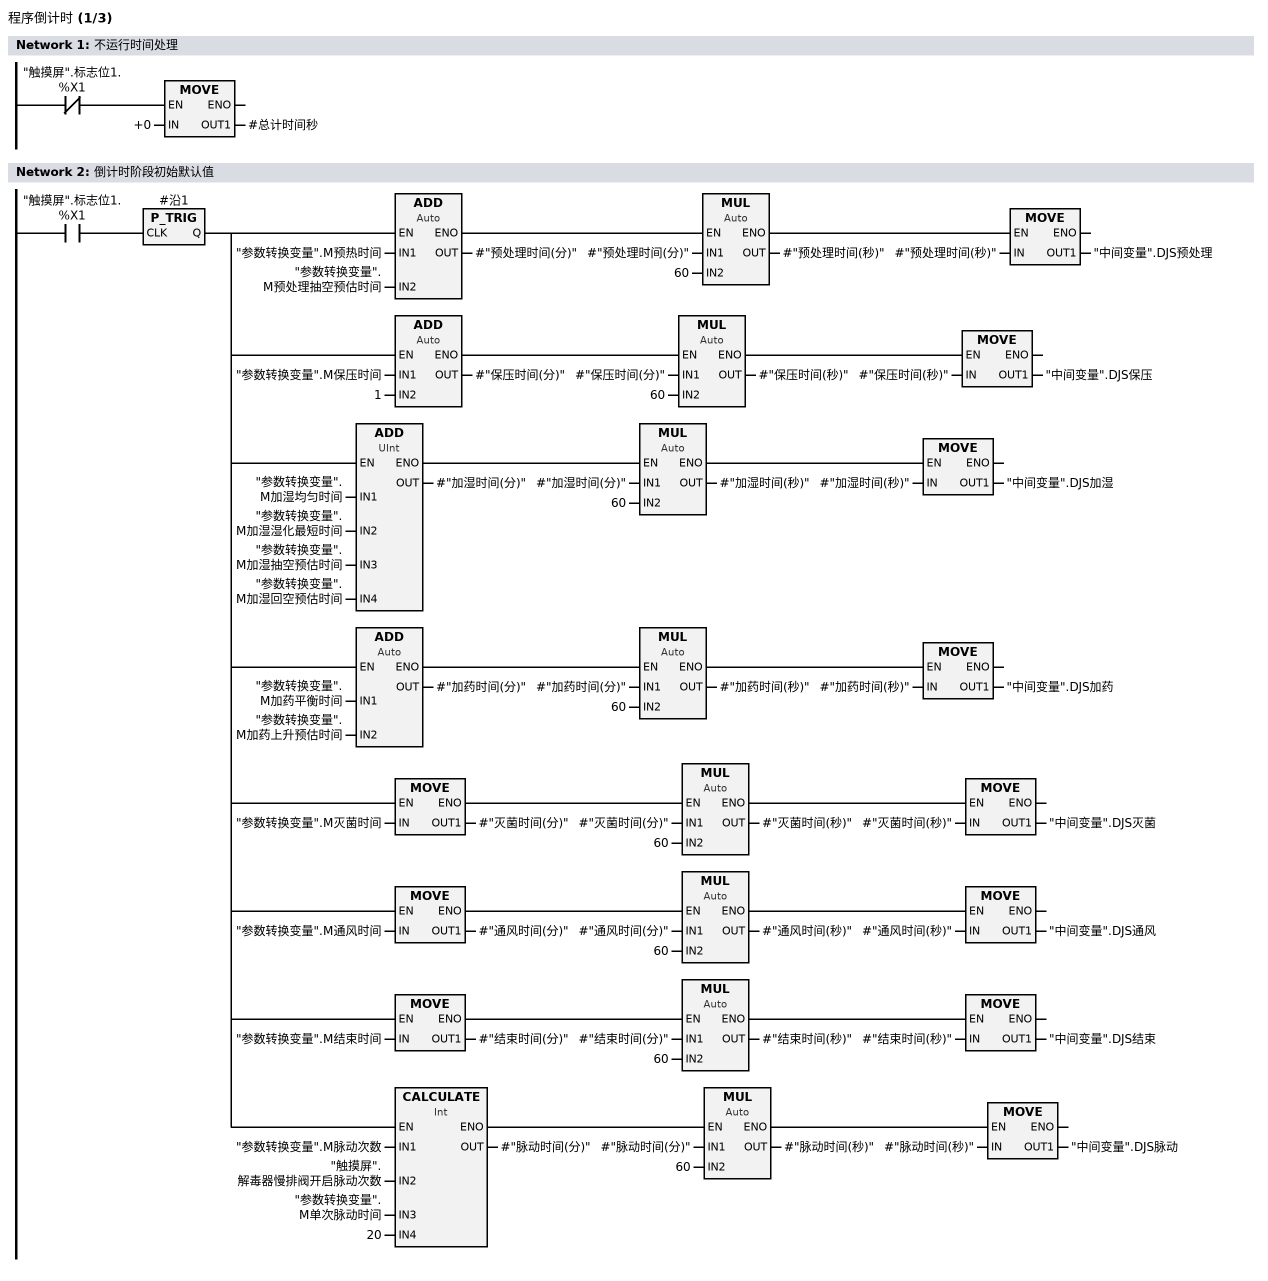
   RUNG wire#powerrail
      I_Contact( "触摸屏".标志位1.%X1 )
      Move(in := +0, out1 => #总计时间秒)
   END_RUNG
   // the same network as SCL:
   IF NOT "触摸屏".标志位1.%X1 THEN #总计时间秒 := +0; END_IF;
END_REGION

REGION Network 2: 倒计时阶段初始默认值
   RUNG wire#powerrail
      Contact( "触摸屏".标志位1.%X1 )
      P_Trig( #沿1 )
      wire#w1
      Add(in1 := "参数转换变量".M预热时间, in2 := "参数转换变量".M预处理抽空预估时间, out => #"预处理时间(分)")
      Mul(in1 := #"预处理时间(分)", in2 := 60, out => #"预处理时间(秒)")
      Move(in := #"预处理时间(秒)", out1 => "中间变量".DJS预处理)
   END_RUNG
   RUNG wire#w1
      Add(in1 := "参数转换变量".M保压时间, in2 := 1, out => #"保压时间(分)")
      Mul(in1 := #"保压时间(分)", in2 := 60, out => #"保压时间(秒)")
      Move(in := #"保压时间(秒)", out1 => "中间变量".DJS保压)
   END_RUNG
   RUNG wire#w1
      { S7_Templates := "SrcType := UInt" } Add(in1 := "参数转换变量".M加湿均匀时间, in2 := "参数转换变量".M加湿湿化最短时间, in3 := "参数转换变量".M加湿抽空预估时间, in4 := "参数转换变量".M加湿回空预估时间, out => #"加湿时间(分)")
      Mul(in1 := #"加湿时间(分)", in2 := 60, out => #"加湿时间(秒)")
      Move(in := #"加湿时间(秒)", out1 => "中间变量".DJS加湿)
   END_RUNG
   RUNG wire#w1
      Add(in1 := "参数转换变量".M加药平衡时间, in2 := "参数转换变量".M加药上升预估时间, out => #"加药时间(分)")
      Mul(in1 := #"加药时间(分)", in2 := 60, out => #"加药时间(秒)")
      Move(in := #"加药时间(秒)", out1 => "中间变量".DJS加药)
   END_RUNG
   RUNG wire#w1
      Move(in := "参数转换变量".M灭菌时间, out1 => #"灭菌时间(分)")
      Mul(in1 := #"灭菌时间(分)", in2 := 60, out => #"灭菌时间(秒)")
      Move(in := #"灭菌时间(秒)", out1 => "中间变量".DJS灭菌)
   END_RUNG
   RUNG wire#w1
      Move(in := "参数转换变量".M通风时间, out1 => #"通风时间(分)")
      Mul(in1 := #"通风时间(分)", in2 := 60, out => #"通风时间(秒)")
      Move(in := #"通风时间(秒)", out1 => "中间变量".DJS通风)
   END_RUNG
   RUNG wire#w1
      Move(in := "参数转换变量".M结束时间, out1 => #"结束时间(分)")
      Mul(in1 := #"结束时间(分)", in2 := 60, out => #"结束时间(秒)")
      Move(in := #"结束时间(秒)", out1 => "中间变量".DJS结束)
   END_RUNG
   RUNG wire#w1
      { S7_Templates := "SrcType := Int"; S7_Expression := "(IN1-IN2)*IN3+IN2*IN4" } Calculate(in1 := "参数转换变量".M脉动次数, in2 := "触摸屏".解毒器慢排阀开启脉动次数, in3 := "参数转换变量".M单次脉动时间, in4 := 20, out => #"脉动时间(分)")
      Mul(in1 := #"脉动时间(分)", in2 := 60, out => #"脉动时间(秒)")
      Move(in := #"脉动时间(秒)", out1 => "中间变量".DJS脉动)
   END_RUNG
   // the same network as SCL:
   #_w1 := "触摸屏".标志位1.%X1 AND NOT #沿1;   // rising edge
   #沿1 := "触摸屏".标志位1.%X1;
   IF #_w1 THEN
       #"预处理时间(分)" := "参数转换变量".M预热时间 + "参数转换变量".M预处理抽空预估时间;
       #"预处理时间(秒)" := #"预处理时间(分)" * 60;
       "中间变量".DJS预处理 := #"预处理时间(秒)";
       #"保压时间(分)" := "参数转换变量".M保压时间 + 1;
       #"保压时间(秒)" := #"保压时间(分)" * 60;
       "中间变量".DJS保压 := #"保压时间(秒)";
       #"加湿时间(分)" := "参数转换变量".M加湿均匀时间 + "参数转换变量".M加湿湿化最短时间 + "参数转换变量".M加湿抽空预估时间 + "参数转换变量".M加湿回空预估时间;
       #"加湿时间(秒)" := #"加湿时间(分)" * 60;
       "中间变量".DJS加湿 := #"加湿时间(秒)";
       #"加药时间(分)" := "参数转换变量".M加药平衡时间 + "参数转换变量".M加药上升预估时间;
       #"加药时间(秒)" := #"加药时间(分)" * 60;
       "中间变量".DJS加药 := #"加药时间(秒)";
       #"灭菌时间(分)" := "参数转换变量".M灭菌时间;
       #"灭菌时间(秒)" := #"灭菌时间(分)" * 60;
       "中间变量".DJS灭菌 := #"灭菌时间(秒)";
       #"通风时间(分)" := "参数转换变量".M通风时间;
       #"通风时间(秒)" := #"通风时间(分)" * 60;
       "中间变量".DJS通风 := #"通风时间(秒)";
       #"结束时间(分)" := "参数转换变量".M结束时间;
       #"结束时间(秒)" := #"结束时间(分)" * 60;
       "中间变量".DJS结束 := #"结束时间(秒)";
       #"脉动时间(分)" := ("参数转换变量".M脉动次数-"触摸屏".解毒器慢排阀开启脉动次数)*"参数转换变量".M单次脉动时间+"触摸屏".解毒器慢排阀开启脉动次数*20;
       #"脉动时间(秒)" := #"脉动时间(分)" * 60;
       "中间变量".DJS脉动 := #"脉动时间(秒)";
   END_IF;
END_REGION

REGION Network 3: 倒计时
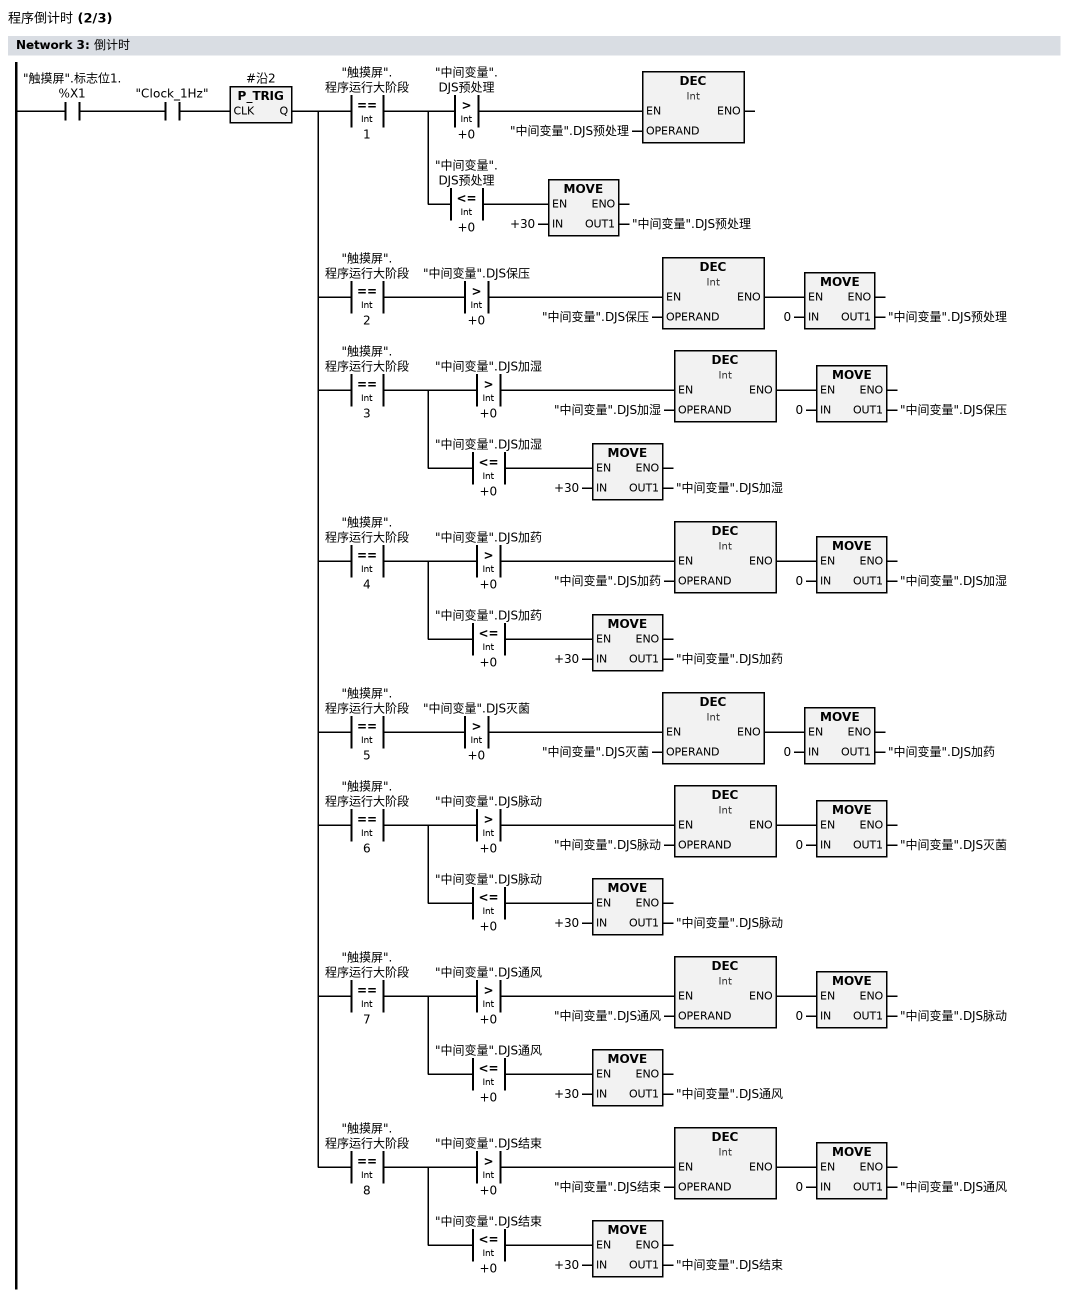
   RUNG wire#powerrail
      Contact( "触摸屏".标志位1.%X1 )
      Contact( "Clock_1Hz" )
      P_Trig( #沿2 )
      wire#w1
      { S7_Templates := "SrcType := Int" } EQ_Contact(in1 := "触摸屏".程序运行大阶段, in2 := 1)
      wire#w2
      { S7_Templates := "SrcType := Int" } GT_Contact(in1 := "中间变量".DJS预处理, in2 := +0)
      { S7_Templates := "DestType := Int" } Dec( "中间变量".DJS预处理 )
   END_RUNG
   RUNG wire#w2
      { S7_Templates := "SrcType := Int" } LE_Contact(in1 := "中间变量".DJS预处理, in2 := +0)
      Move(in := +30, out1 => "中间变量".DJS预处理)
   END_RUNG
   RUNG wire#w1
      { S7_Templates := "SrcType := Int" } EQ_Contact(in1 := "触摸屏".程序运行大阶段, in2 := 2)
      { S7_Templates := "SrcType := Int" } GT_Contact(in1 := "中间变量".DJS保压, in2 := +0)
      { S7_Templates := "DestType := Int" } Dec( "中间变量".DJS保压 )
      Move(in := 0, out1 => "中间变量".DJS预处理)
   END_RUNG
   RUNG wire#w1
      { S7_Templates := "SrcType := Int" } EQ_Contact(in1 := "触摸屏".程序运行大阶段, in2 := 3)
      wire#w3
      { S7_Templates := "SrcType := Int" } GT_Contact(in1 := "中间变量".DJS加湿, in2 := +0)
      { S7_Templates := "DestType := Int" } Dec( "中间变量".DJS加湿 )
      Move(in := 0, out1 => "中间变量".DJS保压)
   END_RUNG
   RUNG wire#w3
      { S7_Templates := "SrcType := Int" } LE_Contact(in1 := "中间变量".DJS加湿, in2 := +0)
      Move(in := +30, out1 => "中间变量".DJS加湿)
   END_RUNG
   RUNG wire#w1
      { S7_Templates := "SrcType := Int" } EQ_Contact(in1 := "触摸屏".程序运行大阶段, in2 := 4)
      wire#w4
      { S7_Templates := "SrcType := Int" } GT_Contact(in1 := "中间变量".DJS加药, in2 := +0)
      { S7_Templates := "DestType := Int" } Dec( "中间变量".DJS加药 )
      Move(in := 0, out1 => "中间变量".DJS加湿)
   END_RUNG
   RUNG wire#w4
      { S7_Templates := "SrcType := Int" } LE_Contact(in1 := "中间变量".DJS加药, in2 := +0)
      Move(in := +30, out1 => "中间变量".DJS加药)
   END_RUNG
   RUNG wire#w1
      { S7_Templates := "SrcType := Int" } EQ_Contact(in1 := "触摸屏".程序运行大阶段, in2 := 5)
      { S7_Templates := "SrcType := Int" } GT_Contact(in1 := "中间变量".DJS灭菌, in2 := +0)
      { S7_Templates := "DestType := Int" } Dec( "中间变量".DJS灭菌 )
      Move(in := 0, out1 => "中间变量".DJS加药)
   END_RUNG
   RUNG wire#w1
      { S7_Templates := "SrcType := Int" } EQ_Contact(in1 := "触摸屏".程序运行大阶段, in2 := 6)
      wire#w5
      { S7_Templates := "SrcType := Int" } GT_Contact(in1 := "中间变量".DJS脉动, in2 := +0)
      { S7_Templates := "DestType := Int" } Dec( "中间变量".DJS脉动 )
      Move(in := 0, out1 => "中间变量".DJS灭菌)
   END_RUNG
   RUNG wire#w5
      { S7_Templates := "SrcType := Int" } LE_Contact(in1 := "中间变量".DJS脉动, in2 := +0)
      Move(in := +30, out1 => "中间变量".DJS脉动)
   END_RUNG
   RUNG wire#w1
      { S7_Templates := "SrcType := Int" } EQ_Contact(in1 := "触摸屏".程序运行大阶段, in2 := 7)
      wire#w6
      { S7_Templates := "SrcType := Int" } GT_Contact(in1 := "中间变量".DJS通风, in2 := +0)
      { S7_Templates := "DestType := Int" } Dec( "中间变量".DJS通风 )
      Move(in := 0, out1 => "中间变量".DJS脉动)
   END_RUNG
   RUNG wire#w6
      { S7_Templates := "SrcType := Int" } LE_Contact(in1 := "中间变量".DJS通风, in2 := +0)
      Move(in := +30, out1 => "中间变量".DJS通风)
   END_RUNG
   RUNG wire#w1
      { S7_Templates := "SrcType := Int" } EQ_Contact(in1 := "触摸屏".程序运行大阶段, in2 := 8)
      wire#w7
      { S7_Templates := "SrcType := Int" } GT_Contact(in1 := "中间变量".DJS结束, in2 := +0)
      { S7_Templates := "DestType := Int" } Dec( "中间变量".DJS结束 )
      Move(in := 0, out1 => "中间变量".DJS通风)
   END_RUNG
   RUNG wire#w7
      { S7_Templates := "SrcType := Int" } LE_Contact(in1 := "中间变量".DJS结束, in2 := +0)
      Move(in := +30, out1 => "中间变量".DJS结束)
   END_RUNG
   // the same network as SCL:
   #_w1 := "触摸屏".标志位1.%X1 AND "Clock_1Hz";
   #_w2 := #_w1 AND NOT #沿2;   // rising edge
   #沿2 := #_w1;
   #_w3 := #_w2 AND ("触摸屏".程序运行大阶段 = 1);
   IF #_w3 AND ("中间变量".DJS预处理 > +0) THEN "中间变量".DJS预处理 := "中间变量".DJS预处理 - 1; END_IF;
   IF #_w3 AND ("中间变量".DJS预处理 <= +0) THEN "中间变量".DJS预处理 := +30; END_IF;
   #_w4 := #_w2 AND ("触摸屏".程序运行大阶段 = 2) AND ("中间变量".DJS保压 > +0);
   IF #_w4 THEN
       "中间变量".DJS保压 := "中间变量".DJS保压 - 1;
       "中间变量".DJS预处理 := 0;
   END_IF;
   #_w5 := #_w2 AND ("触摸屏".程序运行大阶段 = 3);
   #_w6 := #_w5 AND ("中间变量".DJS加湿 > +0);
   IF #_w6 THEN
       "中间变量".DJS加湿 := "中间变量".DJS加湿 - 1;
       "中间变量".DJS保压 := 0;
   END_IF;
   IF #_w5 AND ("中间变量".DJS加湿 <= +0) THEN "中间变量".DJS加湿 := +30; END_IF;
   #_w7 := #_w2 AND ("触摸屏".程序运行大阶段 = 4);
   #_w8 := #_w7 AND ("中间变量".DJS加药 > +0);
   IF #_w8 THEN
       "中间变量".DJS加药 := "中间变量".DJS加药 - 1;
       "中间变量".DJS加湿 := 0;
   END_IF;
   IF #_w7 AND ("中间变量".DJS加药 <= +0) THEN "中间变量".DJS加药 := +30; END_IF;
   #_w9 := #_w2 AND ("触摸屏".程序运行大阶段 = 5) AND ("中间变量".DJS灭菌 > +0);
   IF #_w9 THEN
       "中间变量".DJS灭菌 := "中间变量".DJS灭菌 - 1;
       "中间变量".DJS加药 := 0;
   END_IF;
   #_w10 := #_w2 AND ("触摸屏".程序运行大阶段 = 6);
   #_w11 := #_w10 AND ("中间变量".DJS脉动 > +0);
   IF #_w11 THEN
       "中间变量".DJS脉动 := "中间变量".DJS脉动 - 1;
       "中间变量".DJS灭菌 := 0;
   END_IF;
   IF #_w10 AND ("中间变量".DJS脉动 <= +0) THEN "中间变量".DJS脉动 := +30; END_IF;
   #_w12 := #_w2 AND ("触摸屏".程序运行大阶段 = 7);
   #_w13 := #_w12 AND ("中间变量".DJS通风 > +0);
   IF #_w13 THEN
       "中间变量".DJS通风 := "中间变量".DJS通风 - 1;
       "中间变量".DJS脉动 := 0;
   END_IF;
   IF #_w12 AND ("中间变量".DJS通风 <= +0) THEN "中间变量".DJS通风 := +30; END_IF;
   #_w14 := #_w2 AND ("触摸屏".程序运行大阶段 = 8);
   #_w15 := #_w14 AND ("中间变量".DJS结束 > +0);
   IF #_w15 THEN
       "中间变量".DJS结束 := "中间变量".DJS结束 - 1;
       "中间变量".DJS通风 := 0;
   END_IF;
   IF #_w14 AND ("中间变量".DJS结束 <= +0) THEN "中间变量".DJS结束 := +30; END_IF;
END_REGION

REGION Network 4: 阶段时间累加
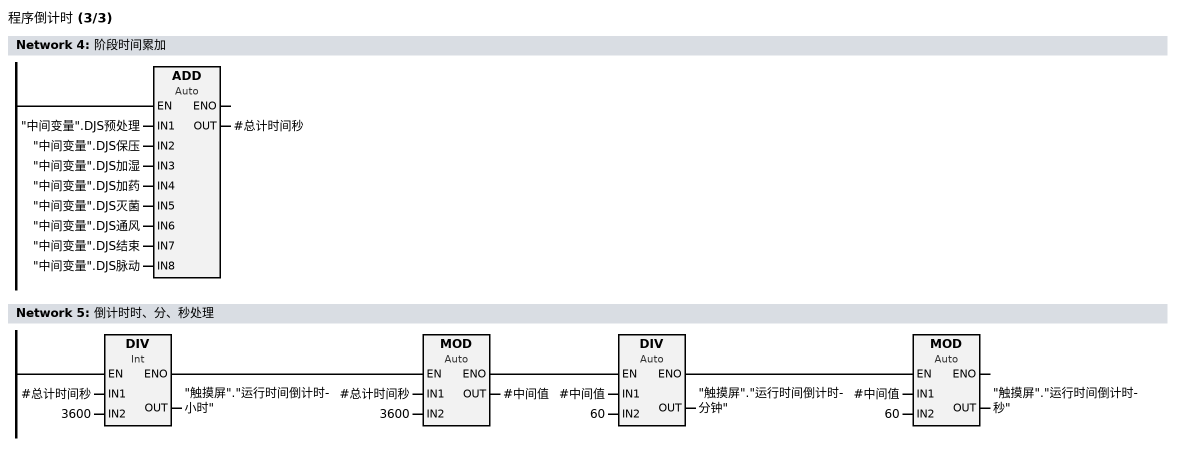
   RUNG wire#powerrail
      Add(in1 := "中间变量".DJS预处理, in2 := "中间变量".DJS保压, in3 := "中间变量".DJS加湿, in4 := "中间变量".DJS加药, in5 := "中间变量".DJS灭菌, in6 := "中间变量".DJS通风, in7 := "中间变量".DJS结束, in8 := "中间变量".DJS脉动, out => #总计时间秒)
   END_RUNG
   // the same network as SCL:
   #总计时间秒 := "中间变量".DJS预处理 + "中间变量".DJS保压 + "中间变量".DJS加湿 + "中间变量".DJS加药 + "中间变量".DJS灭菌 + "中间变量".DJS通风 + "中间变量".DJS结束 + "中间变量".DJS脉动;
END_REGION

REGION Network 5: 倒计时时、分、秒处理
   RUNG wire#powerrail
      { S7_Templates := "SrcType := Int" } Div(in1 := #总计时间秒, in2 := 3600, out => "触摸屏"."运行时间倒计时-小时")
      Mod(in1 := #总计时间秒, in2 := 3600, out => #中间值)
      Div(in1 := #中间值, in2 := 60, out => "触摸屏"."运行时间倒计时-分钟")
      Mod(in1 := #中间值, in2 := 60, out => "触摸屏"."运行时间倒计时-秒")
   END_RUNG
   // the same network as SCL:
   "触摸屏"."运行时间倒计时-小时" := #总计时间秒 / 3600;
   #中间值 := #总计时间秒 MOD 3600;
   "触摸屏"."运行时间倒计时-分钟" := #中间值 / 60;
   "触摸屏"."运行时间倒计时-秒" := #中间值 MOD 60;
END_REGION
END_FUNCTION_BLOCK

FUNCTION "计算倒计时" : Void   // FC6, LAD
{ S7_Optimized_Access := 'TRUE' }
VERSION : 0.1
   VAR_INPUT
      程序运行大阶段 : Int;
   END_VAR
   VAR_OUTPUT
      倒计时总秒数 : DInt;
      各阶段运行时间秒 : DInt;
      循环计数 : Int;
   END_VAR
   VAR_TEMP
      获取当前预制区阶段预估时间秒 : Int;
   END_VAR
BEGIN

REGION Network 1
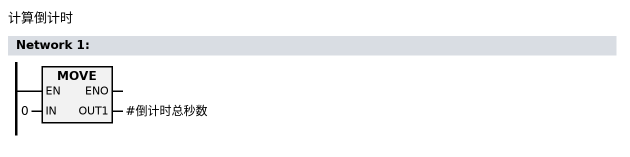
   RUNG wire#powerrail
      Move(in := 0, out1 => #倒计时总秒数)
   END_RUNG
   // the same network as SCL:
   #倒计时总秒数 := 0;
END_REGION

REGION Network 2 (SCL)
   IF #程序运行大阶段 >=0 AND #程序运行大阶段<=10  THEN
       FOR #循环计数 := #程序运行大阶段 TO 10 DO
           IF (#程序运行大阶段 < 8 OR #程序运行大阶段 > 9) THEN

               IF (#循环计数 <> 8 AND #循环计数 <> 9) THEN
                   "获取各阶段预估运行时间秒"(当前阶段名称 := #循环计数,
                                  当前阶段预估时间秒 => #各阶段运行时间秒);
               ELSE
                   #各阶段运行时间秒 := 0;

               END_IF;
           ELSE
               "获取各阶段预估运行时间秒"(当前阶段名称 := #循环计数,
                              当前阶段预估时间秒 => #各阶段运行时间秒);


           END_IF;
           #倒计时总秒数 := #倒计时总秒数 + #各阶段运行时间秒;


       END_FOR;

       END_IF;
END_REGION
END_FUNCTION

FUNCTION "获取各阶段预估运行时间秒" : Void   // FC18, LAD
{ S7_Optimized_Access := 'TRUE' }
VERSION : 0.1
   VAR_INPUT
      当前阶段名称 : Int;
   END_VAR
   VAR_OUTPUT
      当前阶段预估时间秒 : DInt;
   END_VAR
   VAR_TEMP
      沿1 : Bool;
      沿2 : Bool;
   END_VAR
   VAR_TEMP   // added for the SCL form of the ladder/FBD networks
      _w1 : Bool;
   END_VAR
BEGIN

REGION Network 1
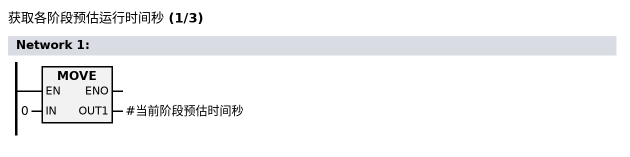
   RUNG wire#powerrail
      Move(in := 0, out1 => #当前阶段预估时间秒)
   END_RUNG
   // the same network as SCL:
   #当前阶段预估时间秒 := 0;
END_REGION

REGION Network 2: 倒计时阶段初始默认值
   // "触摸屏".程序类型.%X2:药罐处理、"触摸屏".程序类型.%X3:泄漏测试
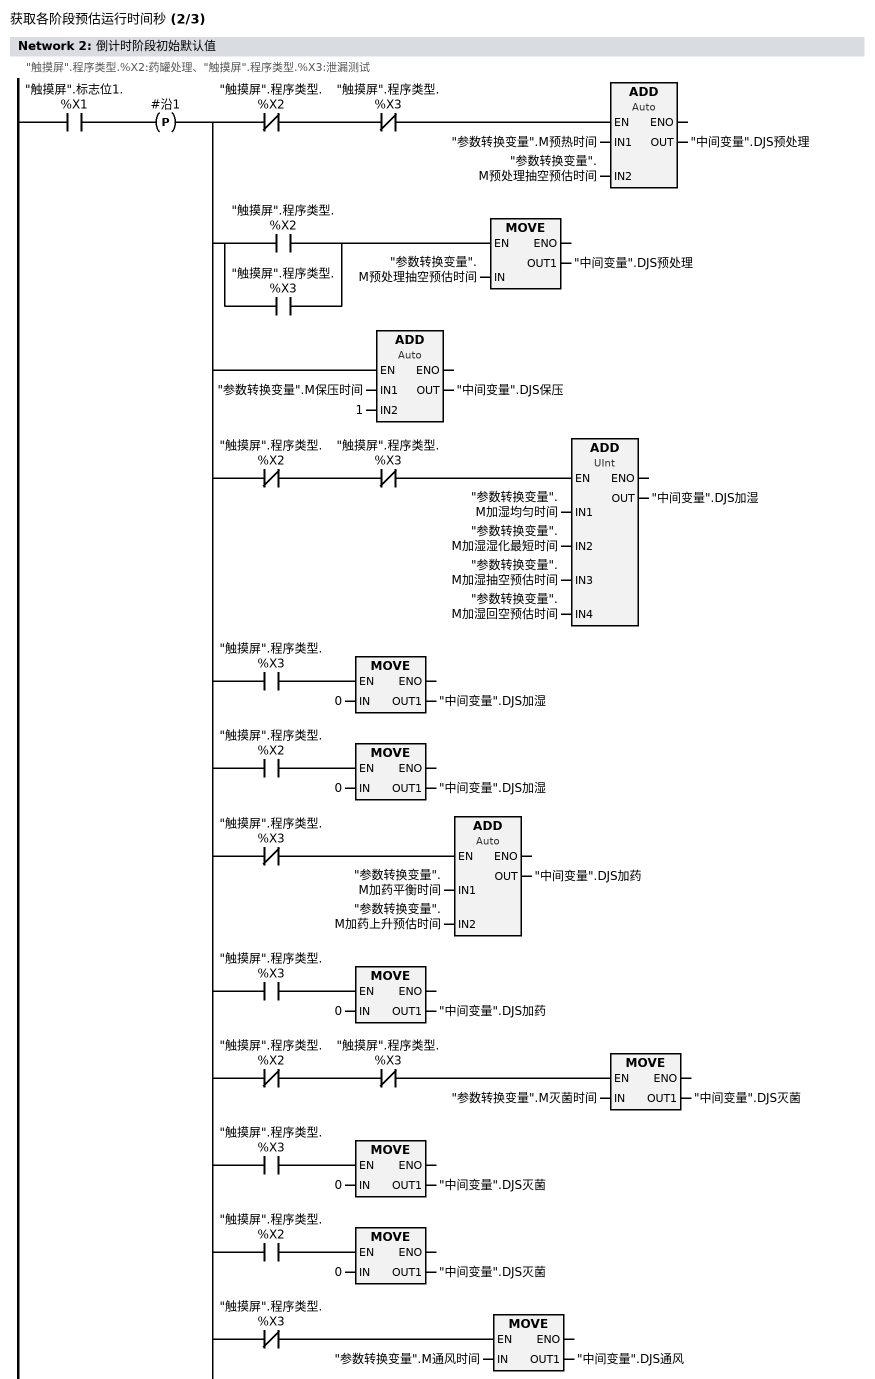
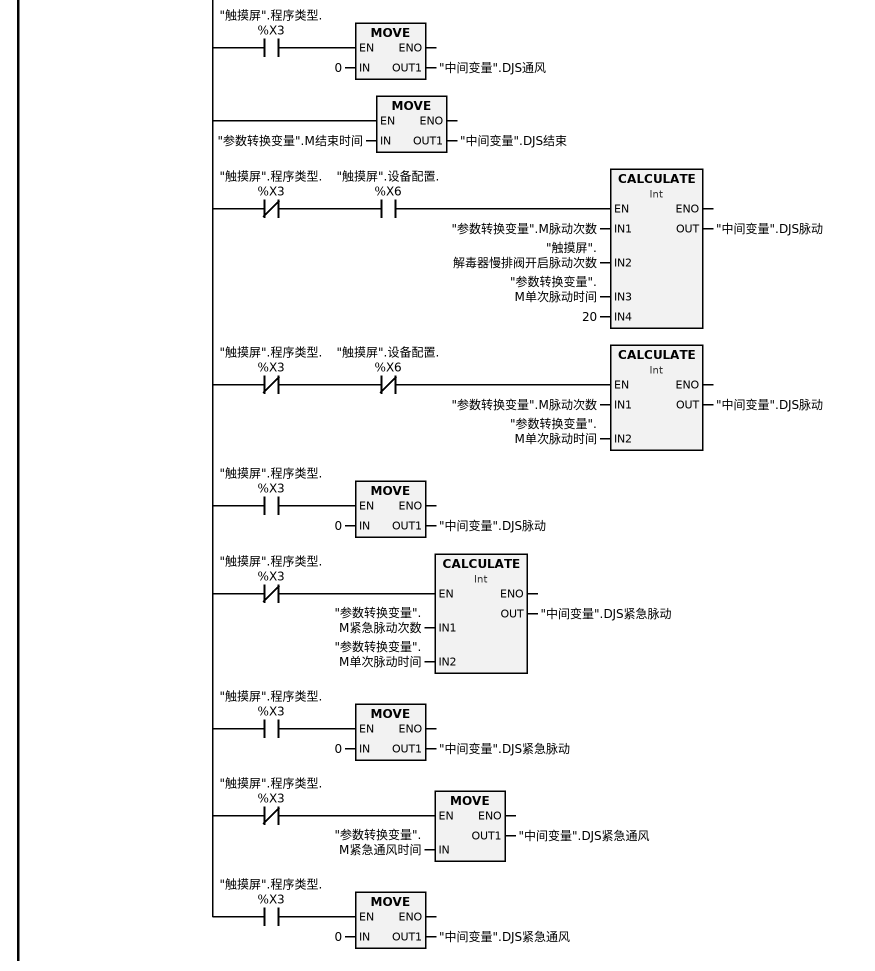
   RUNG wire#powerrail
      Contact( "触摸屏".标志位1.%X1 )
      P_Trig( #沿1 )
      wire#w1
      I_Contact( "触摸屏".程序类型.%X2 )
      I_Contact( "触摸屏".程序类型.%X3 )
      Add(in1 := "参数转换变量".M预热时间, in2 := "参数转换变量".M预处理抽空预估时间, out => "中间变量".DJS预处理)
   END_RUNG
   RUNG wire#w1
      Contact( "触摸屏".程序类型.%X2 )
      wire#w2
      Move(in := "参数转换变量".M预处理抽空预估时间, out1 => "中间变量".DJS预处理)
   END_RUNG
   RUNG wire#w1
      Contact( "触摸屏".程序类型.%X3 )
   END_RUNG wire#w2
   RUNG wire#w1
      Add(in1 := "参数转换变量".M保压时间, in2 := 1, out => "中间变量".DJS保压)
   END_RUNG
   RUNG wire#w1
      I_Contact( "触摸屏".程序类型.%X2 )
      I_Contact( "触摸屏".程序类型.%X3 )
      { S7_Templates := "SrcType := UInt" } Add(in1 := "参数转换变量".M加湿均匀时间, in2 := "参数转换变量".M加湿湿化最短时间, in3 := "参数转换变量".M加湿抽空预估时间, in4 := "参数转换变量".M加湿回空预估时间, out => "中间变量".DJS加湿)
   END_RUNG
   RUNG wire#w1
      Contact( "触摸屏".程序类型.%X3 )
      Move(in := 0, out1 => "中间变量".DJS加湿)
   END_RUNG
   RUNG wire#w1
      Contact( "触摸屏".程序类型.%X2 )
      Move(in := 0, out1 => "中间变量".DJS加湿)
   END_RUNG
   RUNG wire#w1
      I_Contact( "触摸屏".程序类型.%X3 )
      Add(in1 := "参数转换变量".M加药平衡时间, in2 := "参数转换变量".M加药上升预估时间, out => "中间变量".DJS加药)
   END_RUNG
   RUNG wire#w1
      Contact( "触摸屏".程序类型.%X3 )
      Move(in := 0, out1 => "中间变量".DJS加药)
   END_RUNG
   RUNG wire#w1
      I_Contact( "触摸屏".程序类型.%X2 )
      I_Contact( "触摸屏".程序类型.%X3 )
      Move(in := "参数转换变量".M灭菌时间, out1 => "中间变量".DJS灭菌)
   END_RUNG
   RUNG wire#w1
      Contact( "触摸屏".程序类型.%X3 )
      Move(in := 0, out1 => "中间变量".DJS灭菌)
   END_RUNG
   RUNG wire#w1
      Contact( "触摸屏".程序类型.%X2 )
      Move(in := 0, out1 => "中间变量".DJS灭菌)
   END_RUNG
   RUNG wire#w1
      I_Contact( "触摸屏".程序类型.%X3 )
      Move(in := "参数转换变量".M通风时间, out1 => "中间变量".DJS通风)
   END_RUNG
   RUNG wire#w1
      Contact( "触摸屏".程序类型.%X3 )
      Move(in := 0, out1 => "中间变量".DJS通风)
   END_RUNG
   RUNG wire#w1
      Move(in := "参数转换变量".M结束时间, out1 => "中间变量".DJS结束)
   END_RUNG
   RUNG wire#w1
      I_Contact( "触摸屏".程序类型.%X3 )
      Contact( "触摸屏".设备配置.%X6 )
      { S7_Templates := "SrcType := Int"; S7_Expression := "(IN1-IN2)*IN3+IN2*IN4" } Calculate(in1 := "参数转换变量".M脉动次数, in2 := "触摸屏".解毒器慢排阀开启脉动次数, in3 := "参数转换变量".M单次脉动时间, in4 := 20, out => "中间变量".DJS脉动)
   END_RUNG
   RUNG wire#w1
      I_Contact( "触摸屏".程序类型.%X3 )
      I_Contact( "触摸屏".设备配置.%X6 )
      { S7_Templates := "SrcType := Int"; S7_Expression := "IN1*IN2" } Calculate(in1 := "参数转换变量".M脉动次数, in2 := "参数转换变量".M单次脉动时间, out => "中间变量".DJS脉动)
   END_RUNG
   RUNG wire#w1
      Contact( "触摸屏".程序类型.%X3 )
      Move(in := 0, out1 => "中间变量".DJS脉动)
   END_RUNG
   RUNG wire#w1
      I_Contact( "触摸屏".程序类型.%X3 )
      { S7_Templates := "SrcType := Int"; S7_Expression := "IN1*IN2" } Calculate(in1 := "参数转换变量".M紧急脉动次数, in2 := "参数转换变量".M单次脉动时间, out => "中间变量".DJS紧急脉动)
   END_RUNG
   RUNG wire#w1
      Contact( "触摸屏".程序类型.%X3 )
      Move(in := 0, out1 => "中间变量".DJS紧急脉动)
   END_RUNG
   RUNG wire#w1
      I_Contact( "触摸屏".程序类型.%X3 )
      Move(in := "参数转换变量".M紧急通风时间, out1 => "中间变量".DJS紧急通风)
   END_RUNG
   RUNG wire#w1
      Contact( "触摸屏".程序类型.%X3 )
      Move(in := 0, out1 => "中间变量".DJS紧急通风)
   END_RUNG
   // the same network as SCL:
   #_w1 := "触摸屏".标志位1.%X1 AND NOT #沿1;   // rising edge
   #沿1 := "触摸屏".标志位1.%X1;
   IF #_w1 AND NOT "触摸屏".程序类型.%X2 AND NOT "触摸屏".程序类型.%X3 THEN
       "中间变量".DJS预处理 := "参数转换变量".M预热时间 + "参数转换变量".M预处理抽空预估时间;
   END_IF;
   IF #_w1 AND ("触摸屏".程序类型.%X2 OR "触摸屏".程序类型.%X3) THEN "中间变量".DJS预处理 := "参数转换变量".M预处理抽空预估时间; END_IF;
   IF #_w1 THEN "中间变量".DJS保压 := "参数转换变量".M保压时间 + 1; END_IF;
   IF #_w1 AND NOT "触摸屏".程序类型.%X2 AND NOT "触摸屏".程序类型.%X3 THEN
       "中间变量".DJS加湿 := "参数转换变量".M加湿均匀时间 + "参数转换变量".M加湿湿化最短时间 + "参数转换变量".M加湿抽空预估时间 + "参数转换变量".M加湿回空预估时间;
   END_IF;
   IF #_w1 AND "触摸屏".程序类型.%X3 THEN "中间变量".DJS加湿 := 0; END_IF;
   IF #_w1 AND "触摸屏".程序类型.%X2 THEN "中间变量".DJS加湿 := 0; END_IF;
   IF #_w1 AND NOT "触摸屏".程序类型.%X3 THEN "中间变量".DJS加药 := "参数转换变量".M加药平衡时间 + "参数转换变量".M加药上升预估时间; END_IF;
   IF #_w1 AND "触摸屏".程序类型.%X3 THEN "中间变量".DJS加药 := 0; END_IF;
   IF #_w1 AND NOT "触摸屏".程序类型.%X2 AND NOT "触摸屏".程序类型.%X3 THEN "中间变量".DJS灭菌 := "参数转换变量".M灭菌时间; END_IF;
   IF #_w1 AND "触摸屏".程序类型.%X3 THEN "中间变量".DJS灭菌 := 0; END_IF;
   IF #_w1 AND "触摸屏".程序类型.%X2 THEN "中间变量".DJS灭菌 := 0; END_IF;
   IF #_w1 AND NOT "触摸屏".程序类型.%X3 THEN "中间变量".DJS通风 := "参数转换变量".M通风时间; END_IF;
   IF #_w1 AND "触摸屏".程序类型.%X3 THEN "中间变量".DJS通风 := 0; END_IF;
   IF #_w1 THEN "中间变量".DJS结束 := "参数转换变量".M结束时间; END_IF;
   IF #_w1 AND NOT "触摸屏".程序类型.%X3 AND "触摸屏".设备配置.%X6 THEN
       "中间变量".DJS脉动 := ("参数转换变量".M脉动次数-"触摸屏".解毒器慢排阀开启脉动次数)*"参数转换变量".M单次脉动时间+"触摸屏".解毒器慢排阀开启脉动次数*20;
   END_IF;
   IF #_w1 AND NOT "触摸屏".程序类型.%X3 AND NOT "触摸屏".设备配置.%X6 THEN
       "中间变量".DJS脉动 := "参数转换变量".M脉动次数*"参数转换变量".M单次脉动时间;
   END_IF;
   IF #_w1 AND "触摸屏".程序类型.%X3 THEN "中间变量".DJS脉动 := 0; END_IF;
   IF #_w1 AND NOT "触摸屏".程序类型.%X3 THEN "中间变量".DJS紧急脉动 := "参数转换变量".M紧急脉动次数*"参数转换变量".M单次脉动时间; END_IF;
   IF #_w1 AND "触摸屏".程序类型.%X3 THEN "中间变量".DJS紧急脉动 := 0; END_IF;
   IF #_w1 AND NOT "触摸屏".程序类型.%X3 THEN "中间变量".DJS紧急通风 := "参数转换变量".M紧急通风时间; END_IF;
   IF #_w1 AND "触摸屏".程序类型.%X3 THEN "中间变量".DJS紧急通风 := 0; END_IF;
END_REGION

REGION Network 3
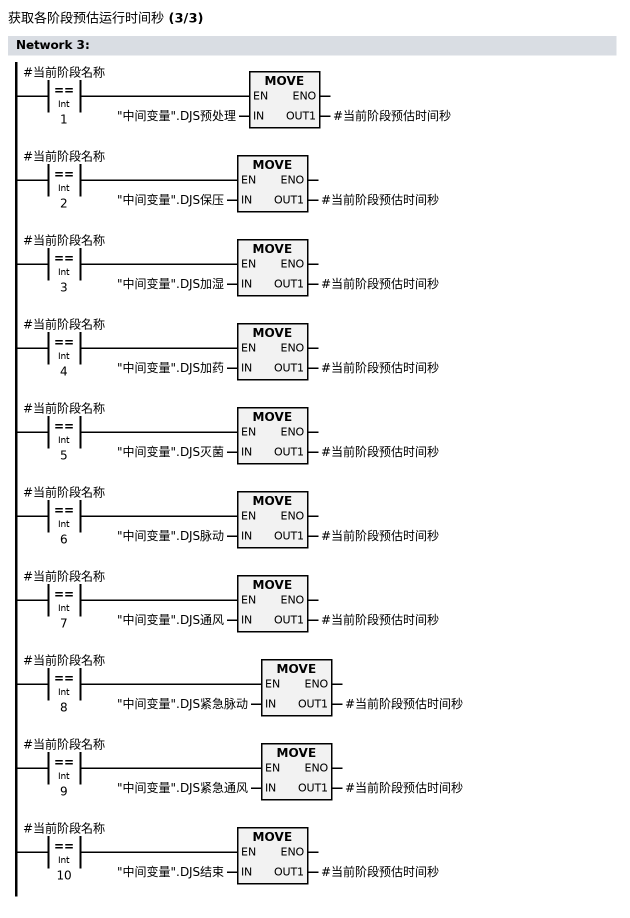
   RUNG wire#powerrail
      { S7_Templates := "SrcType := Int" } EQ_Contact(in1 := #当前阶段名称, in2 := 1)
      Move(in := "中间变量".DJS预处理, out1 => #当前阶段预估时间秒)
   END_RUNG
   RUNG wire#powerrail
      { S7_Templates := "SrcType := Int" } EQ_Contact(in1 := #当前阶段名称, in2 := 2)
      Move(in := "中间变量".DJS保压, out1 => #当前阶段预估时间秒)
   END_RUNG
   RUNG wire#powerrail
      { S7_Templates := "SrcType := Int" } EQ_Contact(in1 := #当前阶段名称, in2 := 3)
      Move(in := "中间变量".DJS加湿, out1 => #当前阶段预估时间秒)
   END_RUNG
   RUNG wire#powerrail
      { S7_Templates := "SrcType := Int" } EQ_Contact(in1 := #当前阶段名称, in2 := 4)
      Move(in := "中间变量".DJS加药, out1 => #当前阶段预估时间秒)
   END_RUNG
   RUNG wire#powerrail
      { S7_Templates := "SrcType := Int" } EQ_Contact(in1 := #当前阶段名称, in2 := 5)
      Move(in := "中间变量".DJS灭菌, out1 => #当前阶段预估时间秒)
   END_RUNG
   RUNG wire#powerrail
      { S7_Templates := "SrcType := Int" } EQ_Contact(in1 := #当前阶段名称, in2 := 6)
      Move(in := "中间变量".DJS脉动, out1 => #当前阶段预估时间秒)
   END_RUNG
   RUNG wire#powerrail
      { S7_Templates := "SrcType := Int" } EQ_Contact(in1 := #当前阶段名称, in2 := 7)
      Move(in := "中间变量".DJS通风, out1 => #当前阶段预估时间秒)
   END_RUNG
   RUNG wire#powerrail
      { S7_Templates := "SrcType := Int" } EQ_Contact(in1 := #当前阶段名称, in2 := 8)
      Move(in := "中间变量".DJS紧急脉动, out1 => #当前阶段预估时间秒)
   END_RUNG
   RUNG wire#powerrail
      { S7_Templates := "SrcType := Int" } EQ_Contact(in1 := #当前阶段名称, in2 := 9)
      Move(in := "中间变量".DJS紧急通风, out1 => #当前阶段预估时间秒)
   END_RUNG
   RUNG wire#powerrail
      { S7_Templates := "SrcType := Int" } EQ_Contact(in1 := #当前阶段名称, in2 := 10)
      Move(in := "中间变量".DJS结束, out1 => #当前阶段预估时间秒)
   END_RUNG
   // the same network as SCL:
   IF #当前阶段名称 = 1 THEN #当前阶段预估时间秒 := "中间变量".DJS预处理; END_IF;
   IF #当前阶段名称 = 2 THEN #当前阶段预估时间秒 := "中间变量".DJS保压; END_IF;
   IF #当前阶段名称 = 3 THEN #当前阶段预估时间秒 := "中间变量".DJS加湿; END_IF;
   IF #当前阶段名称 = 4 THEN #当前阶段预估时间秒 := "中间变量".DJS加药; END_IF;
   IF #当前阶段名称 = 5 THEN #当前阶段预估时间秒 := "中间变量".DJS灭菌; END_IF;
   IF #当前阶段名称 = 6 THEN #当前阶段预估时间秒 := "中间变量".DJS脉动; END_IF;
   IF #当前阶段名称 = 7 THEN #当前阶段预估时间秒 := "中间变量".DJS通风; END_IF;
   IF #当前阶段名称 = 8 THEN #当前阶段预估时间秒 := "中间变量".DJS紧急脉动; END_IF;
   IF #当前阶段名称 = 9 THEN #当前阶段预估时间秒 := "中间变量".DJS紧急通风; END_IF;
   IF #当前阶段名称 = 10 THEN #当前阶段预估时间秒 := "中间变量".DJS结束; END_IF;
END_REGION
END_FUNCTION

// folder: 双泵控制

FUNCTION_BLOCK "双泵控制"   // FB27, LAD
{ S7_Optimized_Access := 'TRUE' }
VERSION : 0.1
   VAR
      双泵配置沿1 : Bool;
      抽空超时报警沿1 : Bool;
      抽空超时报警沿2 : Bool;
      真空泵1过载沿 : Bool;
      真空泵2过载沿 : Bool;
   END_VAR
   VAR_TEMP
      泵编号临时 : Int;
   END_VAR
   VAR_TEMP   // added for the SCL form of the ladder/FBD networks
      _w1 : Bool;
      _w2 : Bool;
      _w3 : Bool;
      _w4 : Bool;
   END_VAR
BEGIN

REGION Network 1: 双泵配置&初始化
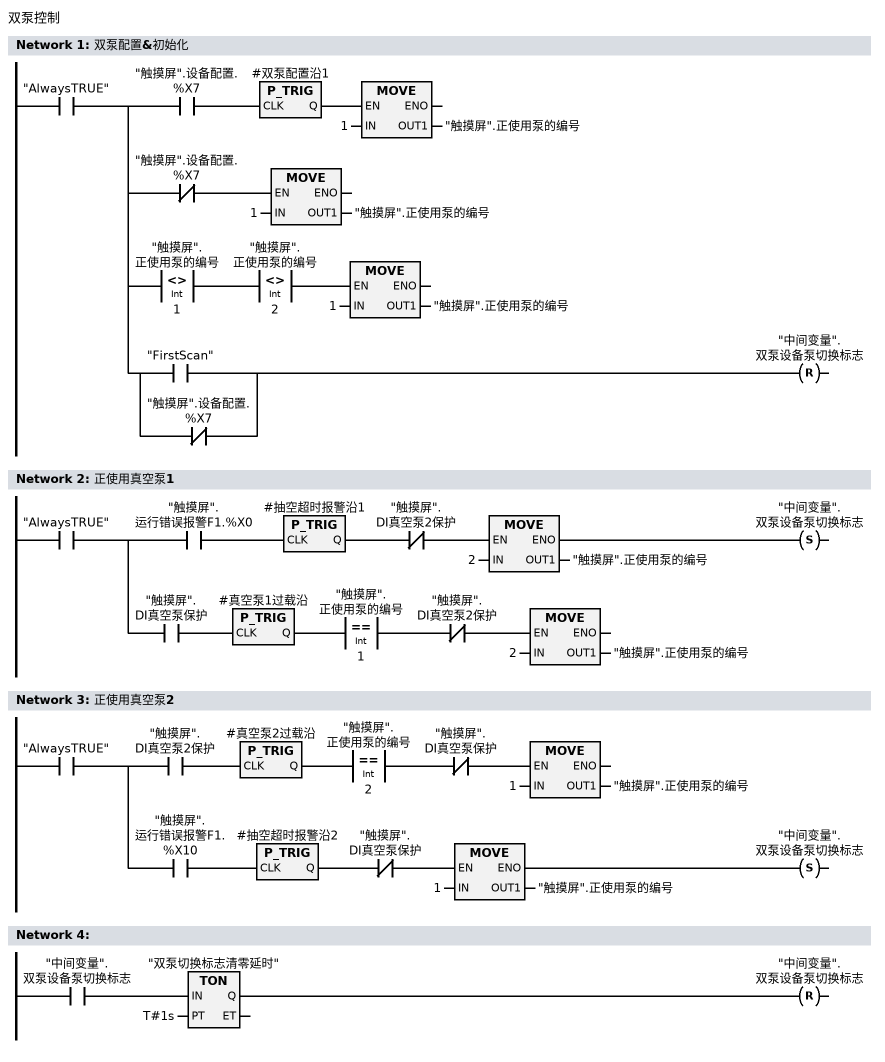
   RUNG wire#powerrail
      Contact( "AlwaysTRUE" )
      wire#w1
      Contact( "触摸屏".设备配置.%X7 )
      P_Trig( #双泵配置沿1 )
      Move(in := 1, out1 => "触摸屏".正使用泵的编号)
   END_RUNG
   RUNG wire#w1
      I_Contact( "触摸屏".设备配置.%X7 )
      Move(in := 1, out1 => "触摸屏".正使用泵的编号)
   END_RUNG
   RUNG wire#w1
      { S7_Templates := "SrcType := Int" } NE_Contact(in1 := "触摸屏".正使用泵的编号, in2 := 1)
      { S7_Templates := "SrcType := Int" } NE_Contact(in1 := "触摸屏".正使用泵的编号, in2 := 2)
      Move(in := 1, out1 => "触摸屏".正使用泵的编号)
   END_RUNG
   RUNG wire#w1
      Contact( "FirstScan" )
      wire#w2
      R_Coil( "中间变量".双泵设备泵切换标志 )
   END_RUNG
   RUNG wire#w1
      I_Contact( "触摸屏".设备配置.%X7 )
   END_RUNG wire#w2
   // the same network as SCL:
   #_w1 := "AlwaysTRUE" AND "触摸屏".设备配置.%X7;
   #_w2 := #_w1 AND NOT #双泵配置沿1;   // rising edge
   #双泵配置沿1 := #_w1;
   IF #_w2 THEN "触摸屏".正使用泵的编号 := 1; END_IF;
   IF "AlwaysTRUE" AND NOT "触摸屏".设备配置.%X7 THEN "触摸屏".正使用泵的编号 := 1; END_IF;
   IF "AlwaysTRUE" AND ("触摸屏".正使用泵的编号 <> 1) AND ("触摸屏".正使用泵的编号 <> 2) THEN "触摸屏".正使用泵的编号 := 1; END_IF;
   IF "AlwaysTRUE" AND ("FirstScan" OR NOT "触摸屏".设备配置.%X7) THEN "中间变量".双泵设备泵切换标志 := FALSE; END_IF;
END_REGION

REGION Network 2: 正使用真空泵1
   RUNG wire#powerrail
      Contact( "AlwaysTRUE" )
      wire#w1
      Contact( "触摸屏".运行错误报警F1.%X0 )
      P_Trig( #抽空超时报警沿1 )
      I_Contact( "触摸屏".DI真空泵2保护 )
      Move(in := 2, out1 => "触摸屏".正使用泵的编号)
      S_Coil( "中间变量".双泵设备泵切换标志 )
   END_RUNG
   RUNG wire#w1
      Contact( "触摸屏".DI真空泵保护 )
      P_Trig( #真空泵1过载沿 )
      { S7_Templates := "SrcType := Int" } EQ_Contact(in1 := "触摸屏".正使用泵的编号, in2 := 1)
      I_Contact( "触摸屏".DI真空泵2保护 )
      Move(in := 2, out1 => "触摸屏".正使用泵的编号)
   END_RUNG
   // the same network as SCL:
   #_w1 := "AlwaysTRUE" AND "触摸屏".运行错误报警F1.%X0;
   #_w2 := #_w1 AND NOT #抽空超时报警沿1;   // rising edge
   #抽空超时报警沿1 := #_w1;
   IF #_w2 AND NOT "触摸屏".DI真空泵2保护 THEN
       "触摸屏".正使用泵的编号 := 2;
       "中间变量".双泵设备泵切换标志 := TRUE;
   END_IF;
   #_w3 := "AlwaysTRUE" AND "触摸屏".DI真空泵保护;
   #_w4 := #_w3 AND NOT #真空泵1过载沿;   // rising edge
   #真空泵1过载沿 := #_w3;
   IF #_w4 AND ("触摸屏".正使用泵的编号 = 1) AND NOT "触摸屏".DI真空泵2保护 THEN "触摸屏".正使用泵的编号 := 2; END_IF;
END_REGION

REGION Network 3: 正使用真空泵2
   RUNG wire#powerrail
      Contact( "AlwaysTRUE" )
      wire#w1
      Contact( "触摸屏".DI真空泵2保护 )
      P_Trig( #真空泵2过载沿 )
      { S7_Templates := "SrcType := Int" } EQ_Contact(in1 := "触摸屏".正使用泵的编号, in2 := 2)
      I_Contact( "触摸屏".DI真空泵保护 )
      Move(in := 1, out1 => "触摸屏".正使用泵的编号)
   END_RUNG
   RUNG wire#w1
      Contact( "触摸屏".运行错误报警F1.%X10 )
      P_Trig( #抽空超时报警沿2 )
      I_Contact( "触摸屏".DI真空泵保护 )
      Move(in := 1, out1 => "触摸屏".正使用泵的编号)
      S_Coil( "中间变量".双泵设备泵切换标志 )
   END_RUNG
   // the same network as SCL:
   #_w1 := "AlwaysTRUE" AND "触摸屏".DI真空泵2保护;
   #_w2 := #_w1 AND NOT #真空泵2过载沿;   // rising edge
   #真空泵2过载沿 := #_w1;
   IF #_w2 AND ("触摸屏".正使用泵的编号 = 2) AND NOT "触摸屏".DI真空泵保护 THEN "触摸屏".正使用泵的编号 := 1; END_IF;
   #_w3 := "AlwaysTRUE" AND "触摸屏".运行错误报警F1.%X10;
   #_w4 := #_w3 AND NOT #抽空超时报警沿2;   // rising edge
   #抽空超时报警沿2 := #_w3;
   IF #_w4 AND NOT "触摸屏".DI真空泵保护 THEN
       "触摸屏".正使用泵的编号 := 1;
       "中间变量".双泵设备泵切换标志 := TRUE;
   END_IF;
END_REGION

REGION Network 4
   "双泵切换标志清零延时".TON(IN := "中间变量".双泵设备泵切换标志, PT := T#1s);
   IF "双泵切换标志清零延时".Q THEN "中间变量".双泵设备泵切换标志 := FALSE; END_IF;
END_REGION
END_FUNCTION_BLOCK